# EPICS autosave request: examples/PSI/lab_setup/plcs_autosave/db/ecmc_test.req
#UPDATE-FREQ=10
#ENABLE-PASS=1
#--------------------------------
# this file contains ASR PVs of the motion controller
# see startup.cmd
#--------------------------------

# Test
$(IOC):Set-Ana-RB
$(IOC):Set-Bin-RB
